// TIA Portal V20 export
Screen "Pop-up_Hmi_Opmodes6_h_Popup"  507x540
  ScreenItem "Background" at 0,0 size 507x540  Type=HmiRectangle
  ScreenItem "Textfeld_1" at 109,102 size 29x30  Type=HmiTextBox
  ScreenItem "Dummy6" at 273,106 size 25x25  Type=HmiRectangle
  ScreenItem "Text_HmiPanelNo" at 136,49 size 160x23  Type=HmiTextBox
  ScreenItem "Descr_OPMode" at 100,26 size 305x20  Type=HmiTextBox
  ScreenItem "Overview_OPMode" at 0,1 size 507x25  Type=HmiTextBox
  ScreenItem "State_OPMode1_Select" at 143,76 size 25x25  Type=HmiTextBox
  ScreenItem "State_OPMode1_NotSelect" at 143,76 size 25x25  Type=HmiTextBox
  ScreenItem "State_OPMode1_Vis" at 143,76 size 25x25  Type=HmiRectangle
  ScreenItem "State_OPMode2_Select" at 169,76 size 25x25  Type=HmiTextBox
  ScreenItem "State_OPMode2_NotSelect" at 169,76 size 25x25  Type=HmiTextBox
  ScreenItem "State_OPMode2_Vis" at 169,76 size 25x25  Type=HmiRectangle
  ScreenItem "State_OPMode3_Select" at 195,76 size 25x25  Type=HmiTextBox
  ScreenItem "State_OPMode3_NotSelect" at 195,76 size 25x25  Type=HmiTextBox
  ScreenItem "State_OPMode3_Vis" at 195,76 size 25x25  Type=HmiRectangle
  ScreenItem "State_OPMode4_Select" at 221,76 size 25x25  Type=HmiTextBox
  ScreenItem "State_OPMode4_NotSelect" at 221,76 size 25x25  Type=HmiTextBox
  ScreenItem "State_OPMode4_Vis" at 221,76 size 25x25  Type=HmiRectangle
  ScreenItem "State_OPMode5_Select" at 247,76 size 25x25  Type=HmiTextBox
  ScreenItem "State_OPMode5_NotSelect" at 247,76 size 25x25  Type=HmiTextBox
  ScreenItem "State_OPMode5_Vis" at 247,76 size 25x25  Type=HmiRectangle
  ScreenItem "State_OPMode6_Select" at 273,76 size 25x25  Type=HmiTextBox
  ScreenItem "State_OPMode6_NotSelect" at 273,76 size 25x25  Type=HmiTextBox
  ScreenItem "State_OPMode6_Vis" at 273,76 size 25x25  Type=HmiRectangle
  ScreenItem "Button_Back" at 1,1 size 90x60  Type=HmiButton
  ScreenItem "Button_Close" at 417,1 size 90x60  Type=HmiButton
  ScreenItem "Text_OPModeArea" at -84,288 size 260x25  Type=HmiTextBox
